// TIA Portal V20 export
// export: Created 2026-10-12T05:42:32.7854364Z, ExportSetting WithDefaults, DisplayName Totally Integrated Automation Portal, DisplayVersion V20, DisplayName TIA Portal Openness, DisplayVersion V20, DisplayName TIA Portal Teamcenter Gateway, DisplayVersion V20, DisplayName TIA Portal Version Control Interface, DisplayVersion V20, DisplayName SINAMICS Startdrive Advanced, DisplayVersion V20 SP1 Update 2, DisplayName SINAMICS Startdrive G110M, G120, G120C, G120D, G120P, G115D, DisplayVersion V20 SP1 Update 2, DisplayName SINAMICS Startdrive G130, G150, S120, S150, SINAMICS MV, G220, S200, S210, DisplayVersion V20 SP1 Update 2, DisplayName STEP 7 Professional, DisplayVersion V20, DisplayName STEP 7 Safety, DisplayVersion V20, DisplayName WinCC Basic/Comfort/Advanced, DisplayVersion V20, DisplayName WinCC Professional, DisplayVersion V20, DisplayName WinCC Unified, DisplayVersion V20
FUNCTION "FRK_SeqCommand" : Bool   // FC134, SCL
{ S7_Optimized_Access := 'TRUE' }
VERSION : 0.1
// stored: AutoNumber true, IsIECCheckEnabled false, SetENOAutomatically false, UDAEnableTagReadback false
   VAR_INPUT
      Value : DInt;
      Label : String;
      Ready : Bool;
      Done : Bool;
      Error : Bool;
      OwnFailure : Bool;
      Diagnostic : "ST_Diagnostic";
   END_VAR
   VAR_IN_OUT
      Seq : "FRK_SequenceCtx";
      Lease : "ST_SequenceCommandLease";
      Execute : Bool;
      Command : DInt;
   END_VAR
   VAR_TEMP
      WaitOk : Bool;
   END_VAR
BEGIN

   #FRK_SeqCommand := FALSE;
   IF NOT #Seq.Running OR #Seq.Error OR #Seq.OwnerIndex <= 0 OR #Seq.ChainIndex <= 0 THEN
       RETURN;
   END_IF;
   IF #Lease.Raised THEN
       IF #Lease.OwnerIndex <> #Seq.OwnerIndex OR #Lease.ChainIndex <> #Seq.ChainIndex OR #Lease.BranchIndex <> #Seq.BranchIndex
           OR #Lease.Step <> #Seq.Step OR #Command <> #Value THEN
           // Another chain owns this command; never borrow its Done result.
           #WaitOk := "FRK_SeqAwait"(Seq := #Seq, Label := 'std.release.commandOwned', Ok := FALSE);
           RETURN;
       END_IF;
       IF #Done THEN
           #FRK_SeqCommand := TRUE;
       ELSIF #Error THEN
           IF #OwnFailure THEN
               #Seq.CommandFailed := TRUE;
               #Seq.HandledDiagnostic := #Diagnostic;
           ELSE
               #Seq.Error := TRUE;
               #Seq.ErrorDiagnostic := #Diagnostic;
           END_IF;
           #Execute := FALSE;
       ELSE
           #WaitOk := "FRK_SeqAwait"(Seq := #Seq, Label := #Label, Ok := FALSE);
       END_IF;
   ELSIF #Ready AND #Lease.ReleasedScan <> #Seq.Scan THEN
       #Lease.OwnerIndex := #Seq.OwnerIndex;
       #Lease.ChainIndex := #Seq.ChainIndex;
       #Lease.BranchIndex := #Seq.BranchIndex;
       #Lease.Step := #Seq.Step;
       #Lease.Raised := TRUE;
       #Seq.CommandIssued := TRUE;
       #Command := #Value;
       #Execute := TRUE;
       #WaitOk := "FRK_SeqAwait"(Seq := #Seq, Label := #Label, Ok := FALSE);
   ELSE
       #WaitOk := "FRK_SeqAwait"(Seq := #Seq, Label := #Label, Ok := FALSE);
   END_IF;
END_FUNCTION
